// TIA Portal V21 export
// export: Created 2026-08-21T20:18:53.8197365Z, ExportSetting None, DisplayName Totally Integrated Automation Portal, DisplayVersion V21, DisplayName STEP 7 Professional, DisplayVersion V21, DisplayName STEP 7 Safety, DisplayVersion V21, DisplayName Tech WebApplication, DisplayVersion V21, DisplayName WinCC Basic/Comfort/Advanced, DisplayVersion V21, DisplayName WinCC Professional, DisplayVersion V21, DisplayName WinCC Unified, DisplayVersion V21
FUNCTION_BLOCK "MTPMonAnaVlv_Type1"   // FB7, FBD
{ S7_Optimized_Access := 'TRUE' }
// stored: MemoryReserve 100, SetENOAutomatically false
   VAR_INPUT
      from_Ctrl { ExternalAccessible := 'False'; ExternalVisible := 'False'; ExternalWritable := 'False'} : "StruCm";
      Service_Occupied { ExternalAccessible := 'False'; ExternalVisible := 'False'; ExternalWritable := 'False'} : Bool;
      Cmd_Auto { ExternalAccessible := 'False'; ExternalVisible := 'False'; ExternalWritable := 'False'} : Bool;
      Cmd_Man { ExternalAccessible := 'False'; ExternalVisible := 'False'; ExternalWritable := 'False'} : Bool;
      Cmd_MVExt { ExternalAccessible := 'False'; ExternalVisible := 'False'; ExternalWritable := 'False'} : Bool;
      Cmd_MVInt { ExternalAccessible := 'False'; ExternalVisible := 'False'; ExternalWritable := 'False'} : Bool;
      Cmd_OpenAut { ExternalAccessible := 'False'; ExternalVisible := 'False'; ExternalWritable := 'False'} : Bool;
      Cmd_CloseAut { ExternalAccessible := 'False'; ExternalVisible := 'False'; ExternalWritable := 'False'} : Bool;
      Cmd_Reset { ExternalAccessible := 'False'; ExternalVisible := 'False'; ExternalWritable := 'False'} : Bool;
      MV_Out_QB { ExternalAccessible := 'False'; ExternalVisible := 'False'; ExternalWritable := 'False'} : Bool := true;
      MV_Unit { ExternalAccessible := 'False'; ExternalVisible := 'False'; ExternalWritable := 'False'} : Int := 1342;
      Intlk04_In01 { ExternalAccessible := 'False'; ExternalVisible := 'False'; ExternalWritable := 'False'} : "DigVal";
      Intlk04_InvIn01 { ExternalAccessible := 'False'; ExternalVisible := 'False'; ExternalWritable := 'False'} : Bool;
      Intlk04_In01String : String;
      Intlk04_In02 { ExternalAccessible := 'False'; ExternalVisible := 'False'; ExternalWritable := 'False'} : "DigVal";
      Intlk04_InvIn02 { ExternalAccessible := 'False'; ExternalVisible := 'False'; ExternalWritable := 'False'} : Bool;
      Intlk04_In02String : String;
      Intlk04_In03 { ExternalAccessible := 'False'; ExternalVisible := 'False'; ExternalWritable := 'False'} : "DigVal";
      Intlk04_InvIn03 { ExternalAccessible := 'False'; ExternalVisible := 'False'; ExternalWritable := 'False'} : Bool;
      Intlk04_In03String : String;
      Intlk04_In04 { ExternalAccessible := 'False'; ExternalVisible := 'False'; ExternalWritable := 'False'} : "DigVal";
      Intlk04_InvIn04 { ExternalAccessible := 'False'; ExternalVisible := 'False'; ExternalWritable := 'False'} : Bool;
      Intlk04_In04String : String;
   END_VAR
   VAR_OUTPUT
      to_ctrl { ExternalAccessible := 'False'; ExternalVisible := 'False'; ExternalWritable := 'False'} : "StruCm";
      MV_Out { ExternalAccessible := 'False'; ExternalVisible := 'False'; ExternalWritable := 'False'} : Word;
      Occupied { ExternalAccessible := 'False'; ExternalVisible := 'False'; ExternalWritable := 'False'} : Bool;   // Occupied by a Service procedure
      AutAct { ExternalAccessible := 'False'; ExternalVisible := 'False'; ExternalWritable := 'False'} : Bool;
      ManAct { ExternalAccessible := 'False'; ExternalVisible := 'False'; ExternalWritable := 'False'} : Bool;
      MV_ExtAct { ExternalAccessible := 'False'; ExternalVisible := 'False'; ExternalWritable := 'False'} : Bool;
      FbkOpenOut { ExternalAccessible := 'False'; ExternalVisible := 'False'; ExternalWritable := 'False'} : Bool;
      FbkCloseOut { ExternalAccessible := 'False'; ExternalVisible := 'False'; ExternalWritable := 'False'} : Bool;
      GrpErr { ExternalAccessible := 'False'; ExternalVisible := 'False'; ExternalWritable := 'False'} : Bool;
   END_VAR
   VAR
      AnOut_IDB { ExternalAccessible := 'False'; ExternalVisible := 'False'; ExternalWritable := 'False'} : "AnOu";
      Intlk04_IDB : "Intlk04";
      VlvAnL_IDB { S7_SetPoint := 'True'} : "VlvAnL";
      MTPMonAnaVlv_IDB { ExternalVisible := 'False'; S7_SetPoint := 'True'} : "MTPMonAnaVlv";
   END_VAR
   VAR_TEMP
      CSF_NOP : "DigVal";
      BadAnIn : "DigVal";
      BadOut : "DigVal";
      Intlock : "DigVal";
   END_VAR
   // Intlk04_In01.Value := true;
   // Intlk04_In02.Value := true;
   // Intlk04_In03.Value := true;
   // Intlk04_In04.Value := true;
BEGIN

REGION Network 1: Convert
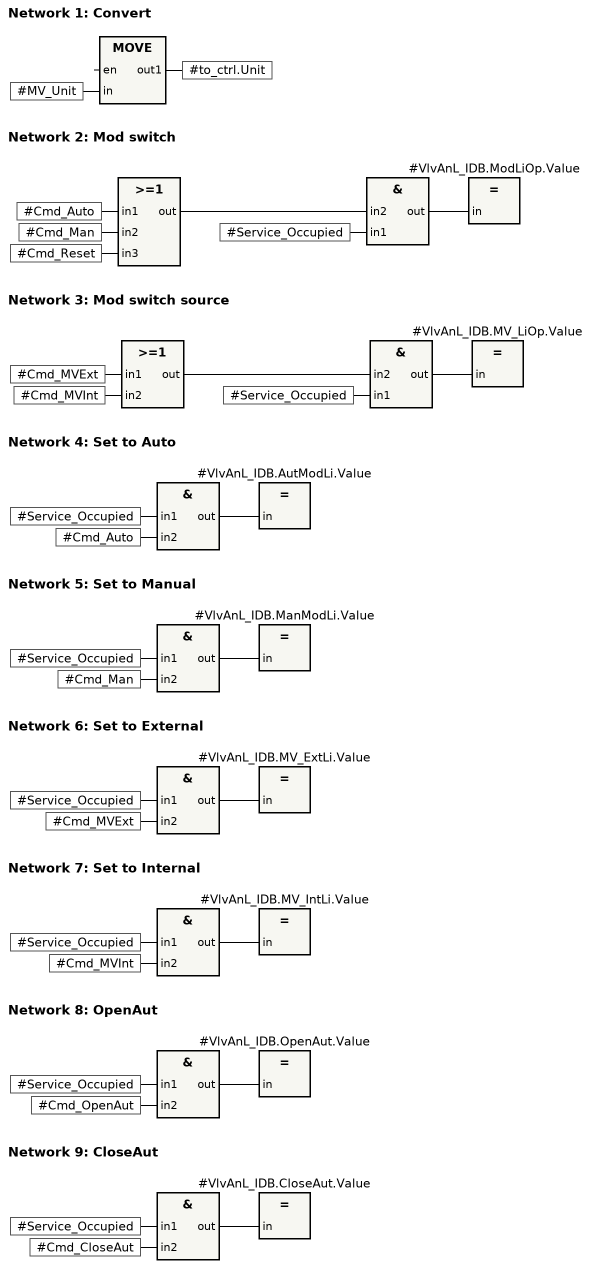
   #to_ctrl.Unit := #MV_Unit;
END_REGION

REGION Network 2: Mod switch
   #VlvAnL_IDB.ModLiOp.Value := (#Cmd_Auto OR #Cmd_Man OR #Cmd_Reset) AND #Service_Occupied;
END_REGION

REGION Network 3: Mod switch source
   #VlvAnL_IDB.MV_LiOp.Value := (#Cmd_MVExt OR #Cmd_MVInt) AND #Service_Occupied;
END_REGION

REGION Network 4: Set to Auto
   #VlvAnL_IDB.AutModLi.Value := #Service_Occupied AND #Cmd_Auto;
END_REGION

REGION Network 5: Set to Manual
   #VlvAnL_IDB.ManModLi.Value := #Service_Occupied AND #Cmd_Man;
END_REGION

REGION Network 6: Set to External
   #VlvAnL_IDB.MV_ExtLi.Value := #Service_Occupied AND #Cmd_MVExt;
END_REGION

REGION Network 7: Set to Internal
   #VlvAnL_IDB.MV_IntLi.Value := #Service_Occupied AND #Cmd_MVInt;
END_REGION

REGION Network 8: OpenAut
   #VlvAnL_IDB.OpenAut.Value := #Service_Occupied AND #Cmd_OpenAut;
END_REGION

REGION Network 9: CloseAut
   #VlvAnL_IDB.CloseAut.Value := #Service_Occupied AND #Cmd_CloseAut;
END_REGION

REGION Network 10: Reset
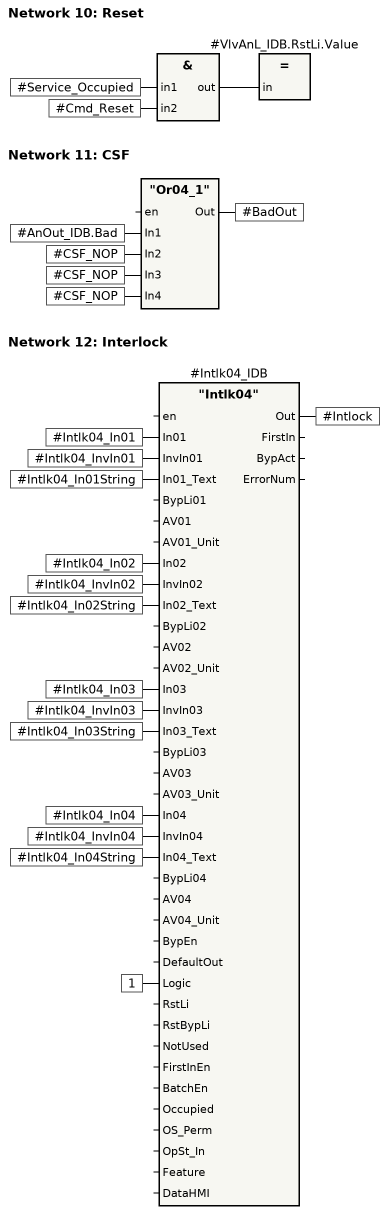
   #VlvAnL_IDB.RstLi.Value := #Service_Occupied AND #Cmd_Reset;
END_REGION

REGION Network 11: CSF
   "Or04_1"(In1 := #AnOut_IDB.Bad, In2 := #CSF_NOP, In3 := #CSF_NOP, In4 := #CSF_NOP, Out => #BadOut);
END_REGION

REGION Network 12: Interlock
   #Intlk04_IDB(In01 := #Intlk04_In01,   // "Intlk04"
                InvIn01 := #Intlk04_InvIn01,
                In01_Text := #Intlk04_In01String,
                In02 := #Intlk04_In02,
                InvIn02 := #Intlk04_InvIn02,
                In02_Text := #Intlk04_In02String,
                In03 := #Intlk04_In03,
                InvIn03 := #Intlk04_InvIn03,
                In03_Text := #Intlk04_In03String,
                In04 := #Intlk04_In04,
                InvIn04 := #Intlk04_InvIn04,
                In04_Text := #Intlk04_In04String,
                Logic := 1,
                Out => #Intlock);
END_REGION

REGION Network 13: VlvAnL
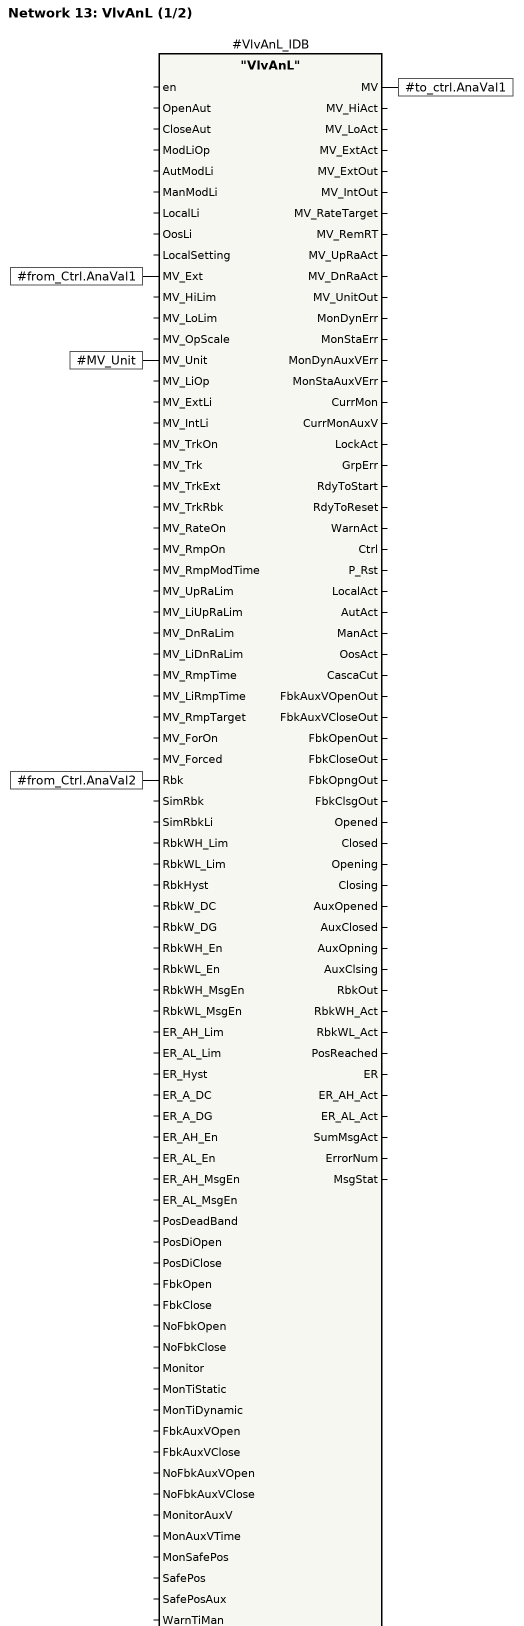
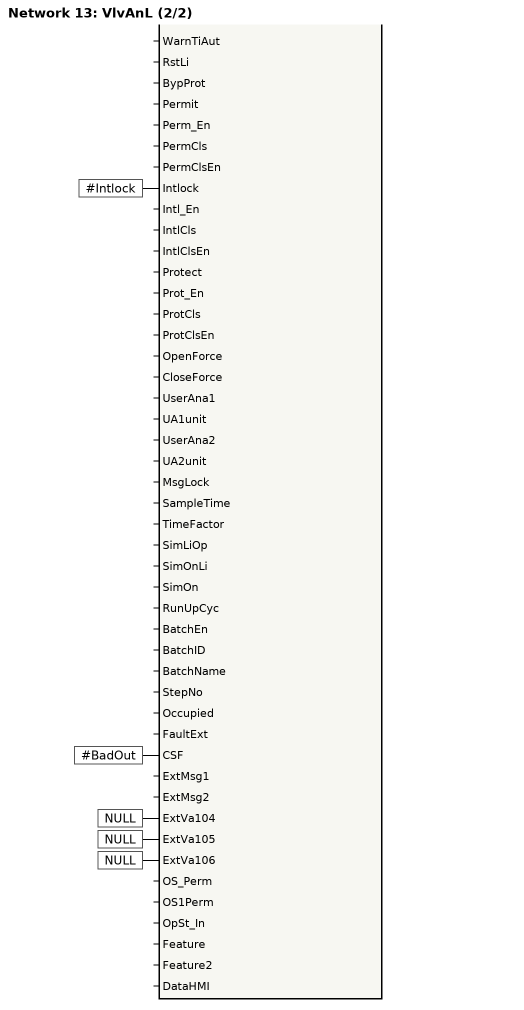
   #VlvAnL_IDB(MV_Ext := #from_Ctrl.AnaVal1,   // "VlvAnL"
               MV_Unit := #MV_Unit,
               Rbk := #from_Ctrl.AnaVal2,
               Intlock := #Intlock,
               CSF := #BadOut,
               ExtVa104 := NULL,
               ExtVa105 := NULL,
               ExtVa106 := NULL,
               MV => #to_ctrl.AnaVal1);
END_REGION

REGION Network 14: Analog Out
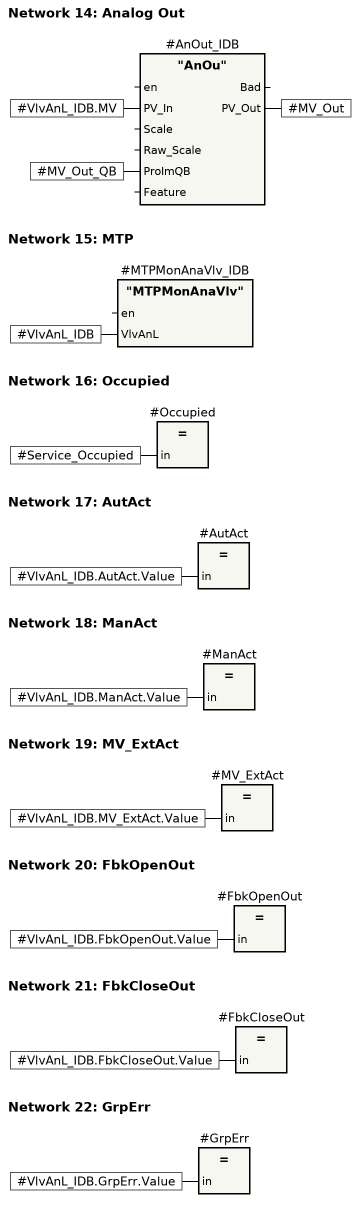
   #AnOut_IDB(PV_In := #VlvAnL_IDB.MV, ProImQB := #MV_Out_QB, PV_Out => #MV_Out);   // "AnOu"
END_REGION

REGION Network 15: MTP
   #MTPMonAnaVlv_IDB(VlvAnL := #VlvAnL_IDB);   // "MTPMonAnaVlv"
END_REGION

REGION Network 16: Occupied
   #Occupied := #Service_Occupied;
END_REGION

REGION Network 17: AutAct
   #AutAct := #VlvAnL_IDB.AutAct.Value;
END_REGION

REGION Network 18: ManAct
   #ManAct := #VlvAnL_IDB.ManAct.Value;
END_REGION

REGION Network 19: MV_ExtAct
   #MV_ExtAct := #VlvAnL_IDB.MV_ExtAct.Value;
END_REGION

REGION Network 20: FbkOpenOut
   #FbkOpenOut := #VlvAnL_IDB.FbkOpenOut.Value;
END_REGION

REGION Network 21: FbkCloseOut
   #FbkCloseOut := #VlvAnL_IDB.FbkCloseOut.Value;
END_REGION

REGION Network 22: GrpErr
   #GrpErr := #VlvAnL_IDB.GrpErr.Value;
END_REGION
END_FUNCTION_BLOCK
